FUNCTION_BLOCK TransferUnit_IMC (* Composite Function Block Type *)
  (* Standard: 61499-2 *)
  (* Version 0.0, 10/23/2026, macie, Schneider Electric, template *)
  PACKAGE Main;
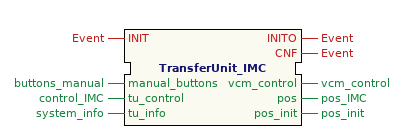
  EVENT_INPUT
    INIT; (* Initialization Request *)
  END_EVENT
  EVENT_OUTPUT
    INITO; (* Initialization Confirm *)
    CNF; (* Execution Confirmation *)
  END_EVENT
  SOCKETS
    manual_buttons : buttons_manual;
    tu_control : control_IMC;
    tu_info : system_info;
  END_SOCKETS
  PLUGS
    vcm_control : vcm_control;
    pos : pos_IMC;
    pos_init : pos_init;
  END_PLUGS
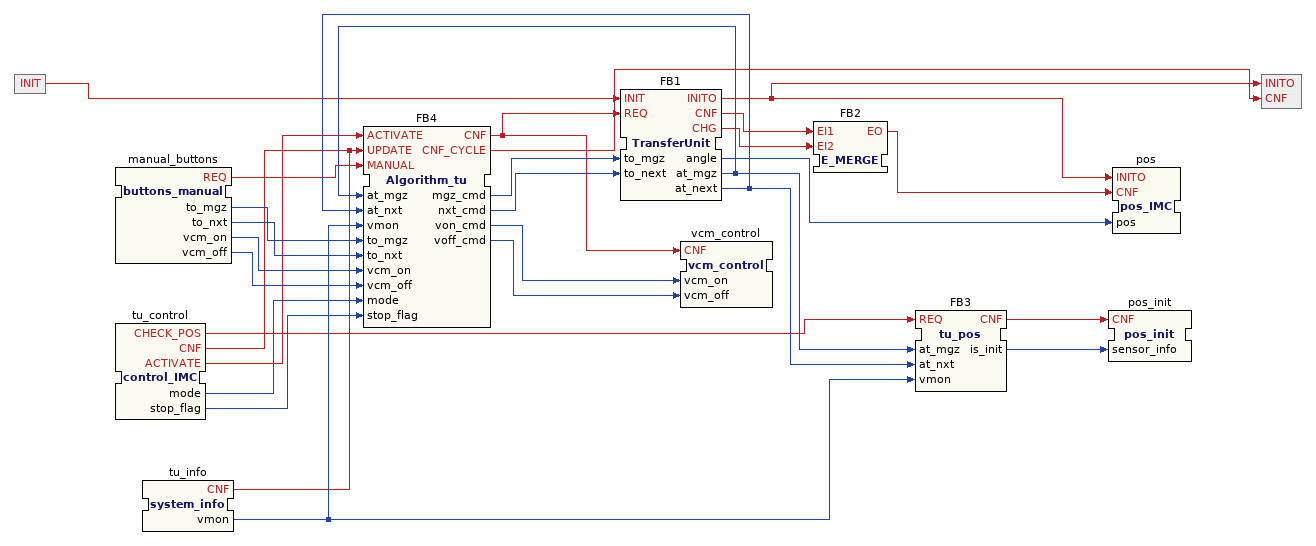
  FBS
    FB1 : TransferUnit;
    FB2 : E_MERGE;
    FB3 : tu_pos;
    FB4 : Algorithm_tu;
  END_FBS
  EVENT_CONNECTIONS
    FB1.INITO TO pos.INITO;
    FB1.CNF TO FB2.EI1;
    FB1.CHG TO FB2.EI2;
    FB2.EO TO pos.CNF;
    INIT TO FB1.INIT;
    FB1.INITO TO INITO;
    tu_control.CHECK_POS TO FB3.REQ;
    manual_buttons.REQ TO FB4.MANUAL;
    tu_control.CNF TO FB4.UPDATE;
    tu_control.ACTIVATE TO FB4.ACTIVATE;
    tu_info.CNF TO FB4.UPDATE;
    FB4.CNF TO FB1.REQ;
    FB4.CNF TO vcm_control.CNF;
    FB3.CNF TO pos_init.CNF;
    FB4.CNF_CYCLE TO CNF;
  END_CONNECTIONS
  DATA_CONNECTIONS
    FB1.angle TO pos.pos;
    FB1.at_mgz TO FB3.at_mgz;
    FB1.at_next TO FB3.at_nxt;
    tu_info.vmon TO FB3.vmon;
    manual_buttons.to_mgz TO FB4.to_mgz;
    manual_buttons.to_nxt TO FB4.to_nxt;
    manual_buttons.vcm_on TO FB4.vcm_on;
    manual_buttons.vcm_off TO FB4.vcm_off;
    tu_control.mode TO FB4.mode;
    tu_control.stop_flag TO FB4.stop_flag;
    tu_info.vmon TO FB4.vmon;
    FB1.at_next TO FB4.at_nxt;
    FB1.at_mgz TO FB4.at_mgz;
    FB4.mgz_cmd TO FB1.to_mgz;
    FB4.nxt_cmd TO FB1.to_next;
    FB4.von_cmd TO vcm_control.vcm_on;
    FB4.voff_cmd TO vcm_control.vcm_off;
    FB3.is_init TO pos_init.sensor_info;
  END_CONNECTIONS
END_FUNCTION_BLOCK
